Fanuc KAREL source: KX00009.KL

PROGRAM KX00009
%NOLOCKGROUP
VAR
  I: INTEGER
  J: INTEGER
  B: BOOLEAN
  F: FILE
  S: STRING[80]
  P: XYZWPR
BEGIN
  STOP
END KX00009
